(* IEC 61131-3 sources: Elmo_Master/Lasal_PRG/MotionTCPDemo/Network, 1 file *)

(* ---- ConfigObjects.st ---- *)
FUNCTION GLOBAL TAB TASK_CONF
_K_TASK, _K_REAL,
_K_END_VAR,

_K_TASK, _K_CYCLIC,
_K_END_VAR,

_K_TASK, _K_BACKGROUND,
_K_END_VAR,

_K_END_CONF
END_FUNCTION

FUNCTION GLOBAL TAB IPR_CONF
_K_IPR
	0$UINT,
_K_END_VAR,
_K_END_CONF
END_FUNCTION

FUNCTION GLOBAL TAB CONFIG_TABLES
00063$UINT,
0$UINT, 1, 59, "_AXISBASE",
0$UINT, 1, 0, "_CHECKSUM",
0$UINT, 0, 5, "_LINKER",
0$UINT, 1, 1, "_LMCABSENCODER",
0$UINT, 1, 123, "_LMCAXIS",
0$UINT, 2, 114, "_LMCAXISBASE",
0$UINT, 1, 33, "_LMCAXISREF",
0$UINT, 1, 43, "_LMCAXISVIS",
0$UINT, 1, 64, "_LMCAXISVISINT",
0$UINT, 1, 1, "_LMCAXISVISLOGHANDLE",
0$UINT, 1, 1, "_LMCAXISVISLOGVIEWER",
0$UINT, 1, 14, "_LMCAXISVISPARA",
0$UINT, 1, 3, "_LMCAXISVOVMONITORING",
0$UINT, 1, 19, "_LMCBASECOORD",
0$UINT, 1, 8, "_LMCBELTAXIS",
0$UINT, 1, 6, "_LMCCALCMODELBASE",
0$UINT, 1, 3, "_LMCCALCMODELCONTROLLER",
0$UINT, 1, 25, "_LMCMATH_SO3",
0$UINT, 1, 76, "_LMCMATHFUNCTIONS",
0$UINT, 1, 1, "_LMCMODULEBASE",
0$UINT, 3, 5, "_LMCPROFILE",
0$UINT, 4, 5, "_LMCPROFILEBASE",
0$UINT, 1, 54, "_LMCPROFILEBUFFER",
0$UINT, 1, 45, "_LMCPROFILELOG",
0$UINT, 1, 31, "_LMCPROFILEVIS",
0$UINT, 1, 21, "_LMCPROFILEVISAXIS",
0$UINT, 1, 42, "_LMCPROFILEVISINT",
0$UINT, 1, 31, "_LMCPROFILEVISMOVEPARA",
0$UINT, 1, 1, "_LMCPUBLISHER",
0$UINT, 1, 12, "_LMCREFBASE",
0$UINT, 2, 23, "_LMCROBOTBASE",
0$UINT, 1, 43, "_LMCROBOTLOG",
0$UINT, 1, 22, "_LMCSAFETY",
0$UINT, 1, 3, "_LMCSPLINEBUFFER",
0$UINT, 1, 24, "_LMCTABLEBUFFER",
0$UINT, 1, 4, "_LMCTOOL",
0$UINT, 1, 1, "_MULTITASK",
0$UINT, 1, 1, "_SIGTCPCOMRECEIVE",
0$UINT, 1, 1, "_SIGTCPDATAMANAGER",
0$UINT, 2, 0, "_STDLIB",
0$UINT, 1, 1, "_TASKOBJECTCONTROL",
0$UINT, 1, 2, "_UDPTRANSCEIVER",
0$UINT, 1, 3, "_UDPTRANSCEIVERINTERFACE",
0$UINT, 1, 48, "CONTROLLER",
0$UINT, 0, 4, "CRITICALSECTION",
0$UINT, 1, 1, "DATAMANAGER",
0$UINT, 1, 1, "DATAMANAGERFIFO",
0$UINT, 1, 0, "DATAMANAGERPRIORITY",
0$UINT, 0, 2, "GETTASKHANDLE",
0$UINT, 1, 0, "MERKER",
0$UINT, 1, 22, "MERKEREX",
0$UINT, 1, 1, "MOVESPLINETABLE",
0$UINT, 1, 1, "RAMRINGBUFFER",
0$UINT, 0, 0, "RECEIVEMSG",
0$UINT, 0, 46, "SIGCLIB",
0$UINT, 1, 11, "STRING",
0$UINT, 1, 86, "STRINGINTERNAL",
0$UINT, 0, 0, "TCP_MOTIONIF_DUMMY",
0$UINT, 1, 20, "TCPCOMMUNICATION",
0$UINT, 1, 0, "TCPCOMMUNICATIONLOGFILTER",
0$UINT, 0, 0, "TCPRT_DATAMANAGER",
0$UINT, 0, 0, "UDPTRANSMISSION",
0$UINT, 1, 3, "VIRTUALBASEINIT",
ONE_CFG$UINT, 0, 0, "ONE_MotionNet",
ONE_CFG$UINT, 0, 0, "ONE_TCPComNet",
ONE_CFG$UINT, 0, 0, "ONE_UDPComNet",
TASK_CFG$UINT, 0, 0, "TASK_CONF",
IPR_CFG$UINT, 0, 0, "IPR_CONF",
PRJ_CFG$UINT, 0, 0, "MotionTCPDemo",
END_FUNCTION

FUNCTION GLOBAL TAB CH_REDIRECT_EMB_TAB
0000$UINT,
00001$UINT,
"TCPCOMMUNICATION;TASKNAME", "\THREADNAME.DATA",
END_FUNCTION
